(* Grating Beam Splitter (GBS): thin ND-framework state-mover wrapper.
   Y mover via FB_PositionStatePMPSND (states OUT, TARGET1a/b, TARGET2a/b,
   TARGET3a/b, TARGET4..6), plus a tick site for two in-beam RTDs gated
   on state. Caller-owned deps injected via FB_Init REFERENCE TO and
   forwarded to fbStates; enum bridge and toggles re-forwarded each cycle. *)
{attribute 'call_after_init'}
FUNCTION_BLOCK FB_GBS
VAR_INPUT
    // Set this to a non-unknown value to request a new move.
    {attribute 'pytmc' := '
        pv: MMS:STATE:SET
        io: io
    '}
    eEnumSet : E_GBS_States;
END_VAR
VAR
    {attribute 'pytmc' := 'pv: RTD:01'}
    fbRTD1 : FB_CC_TempSensor;

    {attribute 'pytmc' := 'pv: RTD:02'}
    fbRTD2 : FB_CC_TempSensor;

    (* REFERENCE TO backing fields populated by FB_Init. Same names as
       FB_Init params; THIS^. disambiguates inside FB_Init.
       Live-bound to caller storage for the lifetime of the FB. *)
    {attribute 'no_copy'}
    aiMotionStage         : REFERENCE TO ARRAY[1..MotionConstants.MAX_STATE_MOTORS] OF I_MotionStage;
    {attribute 'no_copy'}
    astPositionState      : REFERENCE TO ARRAY[1..MotionConstants.MAX_STATE_MOTORS]
                                            OF ARRAY[1..GeneralConstants.MAX_STATES] OF ST_PositionState;
    {attribute 'no_copy'}
    fbFFHWO               : REFERENCE TO FB_HardwareFFOutput;
    {attribute 'no_copy'}
    fbArbiter             : REFERENCE TO FB_Arbiter;
    sDeviceName           : STRING;
    sTransitionKey        : STRING;
    bEnableMotion         : BOOL := TRUE;
    bEnableBeamParams     : BOOL;
    bEnablePositionLimits : BOOL;
    bReadDBNow            : BOOL;
    bFileReaderBusy       : REFERENCE TO BOOL;
    bFileReaderError      : REFERENCE TO BOOL;

    (* One configurator per GBS state (OUT + 9 targets). Writes the
       per-state sName and fDelta. Ticked cyclically in the body AFTER
       fbStates so its writes win over the template baseline
       FB_StateSetup applied via FB_CC_StatePMPSConfig. Idempotent once
       stPositionState.bUpdated trips. *)
    afbStateDefaults : ARRAY[1..10] OF FB_CC_InternalStateConfig[
        (stPositionState := astPositionState[1][E_GBS_States.OUT],
         sName           := 'OUT',
         fDelta          := FDELTA_DEFAULT),
        (stPositionState := astPositionState[1][E_GBS_States.TARGET1a],
         sName           := 'TARGET1a',
         fDelta          := FDELTA_DEFAULT),
        (stPositionState := astPositionState[1][E_GBS_States.TARGET1b],
         sName           := 'TARGET1b',
         fDelta          := FDELTA_DEFAULT),
        (stPositionState := astPositionState[1][E_GBS_States.TARGET2a],
         sName           := 'TARGET2a',
         fDelta          := FDELTA_DEFAULT),
        (stPositionState := astPositionState[1][E_GBS_States.TARGET2b],
         sName           := 'TARGET2b',
         fDelta          := FDELTA_DEFAULT),
        (stPositionState := astPositionState[1][E_GBS_States.TARGET3a],
         sName           := 'TARGET3a',
         fDelta          := FDELTA_DEFAULT),
        (stPositionState := astPositionState[1][E_GBS_States.TARGET3b],
         sName           := 'TARGET3b',
         fDelta          := FDELTA_DEFAULT),
        (stPositionState := astPositionState[1][E_GBS_States.TARGET4],
         sName           := 'TARGET4',
         fDelta          := FDELTA_DEFAULT),
        (stPositionState := astPositionState[1][E_GBS_States.TARGET5],
         sName           := 'TARGET5',
         fDelta          := FDELTA_DEFAULT),
        (stPositionState := astPositionState[1][E_GBS_States.TARGET6],
         sName           := 'TARGET6',
         fDelta          := FDELTA_DEFAULT)
    ];

    {attribute 'pytmc' := 'pv: MMS'}
    fbStates : FB_PositionStatePMPSND(
        aiMotionStage         := aiMotionStage,
        astPositionState      := astPositionState,
        nActiveMotorCount     := 1,
        eEnumSet              := eEnumSet,
        eEnumGet              := eEnumGet,
        bEnableMotion         := bEnableMotion,
        eMotionRequestPolicy  := E_MotionRequestPolicy.INTERRUPT,
        bEnableBeamParams     := bEnableBeamParams,
        bEnablePositionLimits := bEnablePositionLimits,
        bReadDBNow            := bReadDBNow,
        bFileReaderBusy       := bFileReaderBusy,
        bFileReaderError      := bFileReaderError,
        fbFFHWO               := fbFFHWO,
        fbArbiter             := fbArbiter,
        sDeviceName           := sDeviceName,
        sTransitionKey        := sTransitionKey
    );
    i : UINT;
END_VAR
VAR_OUTPUT
    // The current position state as an enum.
    {attribute 'pytmc' := '
        pv: MMS:STATE:GET
        io: i
    '}
    eEnumGet: E_GBS_States;
    // The PMPS database lookup associated with the current position state.
    stDbStateParams: ST_DbStateParams;
END_VAR
VAR CONSTANT
    (* GBS-wide default tolerance for state in-position detection,
       applied per-state by afbStateDefaults. *)
    FDELTA_DEFAULT : LREAL := 2;
END_VAR

(* Nil-ref guards: every REFERENCE TO backing field must be bound. *)
IF NOT __ISVALIDREF(aiMotionStage)
   OR NOT __ISVALIDREF(astPositionState)
   OR NOT __ISVALIDREF(fbFFHWO)
   OR NOT __ISVALIDREF(fbArbiter) THEN
    RETURN;
END_IF

(* Device-side per-state defaults (afbStateDefaults) are written
   once in FB_CC_InternalStateConfig.CallAfterInit; no cyclic tick. *)
fbStates(stDbStateParams=> stDbStateParams);

(* In-beam RTDs: only fault when something is actually in the beam
   (i.e. not OUT). Driven by the PMPS DB temp setpoint. *)
fbRTD1(
    fFaultThreshold := fbStates.stDbStateParams.stReactiveParams.nTempSP,
    bVeto           := eEnumGet = E_GBS_States.OUT,
    sDevName        := sDeviceName,
    io_fbFFHWO      := fbFFHWO
);
fbRTD2(
    fFaultThreshold := fbStates.stDbStateParams.stReactiveParams.nTempSP,
    bVeto           := eEnumGet = E_GBS_States.OUT,
    sDevName        := sDeviceName,
    io_fbFFHWO      := fbFFHWO
);

(* Auto-fired after FB_Init. fbStates' inline-init ran first and
   forwarded nil refs, so this re-supplies the now-valid refs via
   fbStates.CallAfterInitStateMover / CallAfterInitPMPS and writes the
   per-state device defaults. *)
{attribute 'call_after_init'}
METHOD CallAfterInit
afbStateDefaults[1].CallAfterInit(stPositionState := THIS^.astPositionState[1][E_GBS_States.OUT]);
afbStateDefaults[2].CallAfterInit(stPositionState := THIS^.astPositionState[1][E_GBS_States.TARGET1a]);
afbStateDefaults[3].CallAfterInit(stPositionState := THIS^.astPositionState[1][E_GBS_States.TARGET1b]);
afbStateDefaults[4].CallAfterInit(stPositionState := THIS^.astPositionState[1][E_GBS_States.TARGET2a]);
afbStateDefaults[5].CallAfterInit(stPositionState := THIS^.astPositionState[1][E_GBS_States.TARGET2b]);
afbStateDefaults[6].CallAfterInit(stPositionState := THIS^.astPositionState[1][E_GBS_States.TARGET3a]);
afbStateDefaults[7].CallAfterInit(stPositionState := THIS^.astPositionState[1][E_GBS_States.TARGET3b]);
afbStateDefaults[8].CallAfterInit(stPositionState := THIS^.astPositionState[1][E_GBS_States.TARGET4]);
afbStateDefaults[9].CallAfterInit(stPositionState := THIS^.astPositionState[1][E_GBS_States.TARGET5]);
afbStateDefaults[10].CallAfterInit(stPositionState := THIS^.astPositionState[1][E_GBS_States.TARGET6]);

THIS^.fbStates.CallAfterInitStateMover(
    aiMotionStage         := aiMotionStage,
    astPositionState      := astPositionState,
    nActiveMotorCount     := 1,
    eEnumSet              := eEnumSet,
    eEnumGet              := eEnumGet,
    bEnableMotion         := bEnableMotion,
    eMotionRequestPolicy  := E_MotionRequestPolicy.INTERRUPT,
);

THIS^.fbStates.CallAfterInitPMPS(
    aiMotionStage         := aiMotionStage,
    astPositionState      := astPositionState,
    bEnableBeamParams     := bEnableBeamParams,
    bEnablePositionLimits := bEnablePositionLimits,
    bReadDBNow            := bReadDBNow,
    bFileReaderBusy       := bFileReaderBusy,
    bFileReaderError      := bFileReaderError,
    fbFFHWO               := fbFFHWO,
    fbArbiter             := fbArbiter,
    sDeviceName           := sDeviceName,
    sTransitionKey        := sTransitionKey
);
END_METHOD

(* Stores FB_Init inputs into instance fields; every non-value input is
   REFERENCE TO, REF= bound for the FB lifetime. fbStates inline-init
   captured these params at construction, so this records the same refs
   on THIS^ for body use and live caller writes. *)
{attribute 'analysis' := '-33'}
METHOD FB_Init : BOOL
VAR_INPUT
    bInitRetains           : BOOL;
    bInCopyCode            : BOOL;
    aiMotionStage          : REFERENCE TO ARRAY[1..MotionConstants.MAX_STATE_MOTORS] OF I_MotionStage;
    astPositionState       : REFERENCE TO ARRAY[1..MotionConstants.MAX_STATE_MOTORS]
                                            OF ARRAY[1..GeneralConstants.MAX_STATES] OF ST_PositionState;
    fbFFHWO                : REFERENCE TO FB_HardwareFFOutput;
    fbArbiter              : REFERENCE TO FB_Arbiter;
    sDeviceName            : STRING;
    sTransitionKey         : STRING;
    bEnableBeamParams      : BOOL;
    bEnablePositionLimits  : BOOL;
    bReadDBNow             : BOOL;
    bFileReaderBusy       : REFERENCE TO BOOL;
    bFileReaderError      : REFERENCE TO BOOL;
END_VAR
THIS^.aiMotionStage    REF= aiMotionStage;
THIS^.astPositionState REF= astPositionState;
THIS^.fbFFHWO          REF= fbFFHWO;
THIS^.fbArbiter        REF= fbArbiter;
THIS^.sDeviceName      := sDeviceName;
THIS^.sTransitionKey   := sTransitionKey;
THIS^.bEnableBeamParams     := bEnableBeamParams;
THIS^.bEnablePositionLimits := bEnablePositionLimits;
THIS^.bReadDBNow            := bReadDBNow;
THIS^.bFileReaderBusy       REF= bFileReaderBusy;
THIS^.bFileReaderError      REF= bFileReaderError;
END_METHOD

END_FUNCTION_BLOCK

(* stored: Version 1.1.0.1
   POU FB_GBS: Id {0c826496-bbe5-4d0f-95cc-b97d4fbafab2}, SpecialFunc None
   Method CallAfterInit: Id {0c826497-bbe5-4d0f-95cc-b97d4fbafab3}
   Method FB_init: Id {0c826498-bbe5-4d0f-95cc-b97d4fbafab4} *)
